(*
SPDX-FileCopyrightText: c 2026 Oleksandr Tiutyk <trofimich@gmail.com>
SPDX-License-Identifier: MIT
License: https://opensource.org/license/mit
*)

(*!
<summary>Checks release of populated storage and fresh allocation on reuse.</summary>
<description>
Owns a list and its copied entries. Use from one task at a stable address.
Teardown clears surviving entries before publication.
</description>
*)

{attribute 'no_assign'}
{attribute 'no_explicit_call' := 'do not call this function block directly'}
FUNCTION_BLOCK DynamicListClearTest EXTENDS TOF_Testing.SingleCycleTest
VAR_STAT
	{attribute 'hide'}
	_ClassName : STRING := __POUNAME();
END_VAR
VAR
	_List : TOF_Collections.List<0>(valueValidator := 0);
END_VAR

(*!
<summary>Checks release of populated storage and fresh allocation on reuse.</summary>
*)
METHOD PROTECTED ExecuteTest
VAR
	values : ARRAY [0..5] OF STRING := ['String0', 'String1', 'String2', 'String3', 'String4', 'String5'];
END_VAR
_List.AppendCopy(value := values[0]);
_List.AppendCopy(value := values[1]);
_List.AppendCopy(value := values[2]);
_List.AppendCopy(value := values[3]);
_List.AppendCopy(value := values[4]);
_List.AppendCopy(value := values[5]);

Assert.ThatBool(
	actual := _List.Length = 6 AND_THEN _List.Capacity >= 6,
	message := "Clear fixture must contain six live entries"
).IsTrue();

_List.Clear();

Assert.ThatBool(
	actual := _List.Empty AND_THEN _List.Length = 0 AND_THEN _List.Capacity = 0,
	message := "Clear must empty the dynamic list and release its capacity"
).IsTrue();

_List.AppendCopy(value := values[5]);

Assert.ThatBool(
	actual := _List.Length = 1 AND_THEN _List.Get(index := 0).AsString255() = 'String5',
	message := "The cleared list must accept a fresh value"
).IsTrue();
END_METHOD

(*!
<summary>Clears the fixture before the runner publishes the result.</summary>
<description>
Also runs after an unexpected exception interrupts the case.
</description>
*)
METHOD PROTECTED AfterTest
_List.Clear();
END_METHOD

//! <summary>Borrows the concrete class name. Callers must not modify it.</summary>
{attribute 'monitoring' := 'call'}
PROPERTY ClassName : REFERENCE TO STRING
GET
ClassName REF= _ClassName;
END_GET
END_PROPERTY

//! <summary>Borrows the compiler-initialized namespace name. Callers must not modify it.</summary>
{attribute 'monitoring' := 'call'}
PROPERTY NamespaceName : REFERENCE TO STRING
GET
NamespaceName REF= CurrentNamespace.Name;
END_GET
END_PROPERTY

//! <summary>Reports the concrete instance size in bytes.</summary>
{attribute 'monitoring' := 'call'}
PROPERTY SelfSize : ULINT
GET
SelfSize := XSIZEOF(THIS^);
END_GET
END_PROPERTY

END_FUNCTION_BLOCK

(* stored: Version 1.1.0.1
   POU DynamicListClearTest: Id {4bfc7e56-b24a-4a5e-87fb-d1885d23bb9b}, SpecialFunc None
   Method ExecuteTest: Id {9294a094-db16-493f-8629-acebfd4257b6}
   Method AfterTest: Id {449239a7-b620-4796-8be3-f33d80e26b3e}
   Property ClassName: Id {6b4de815-251f-404f-a085-0b24fa36e2ef}
   Get Get: Id {80fb716f-f022-4375-a4c7-4f12b19ff911}
   Property NamespaceName: Id {16bab229-1cec-4012-b352-b05624dd032d}
   Get Get: Id {f726c8d1-1e84-4453-b710-1dee4708deea}
   Property SelfSize: Id {12cbab9f-8e2e-482d-989b-99cb3bb0ca75}
   Get Get: Id {e0a92779-d1f1-4385-a7e1-008ec68132c4} *)
